Fanuc KAREL source: kd00041.KL

-- PROVISIONAL review KL for V940-1; original PC SHA256 db74242f19a3847c4d94c9fab1e78f44e8e95f5fcd8958c4a07cd94807cec2c1
-- Incomplete behavior may be omitted. Consult companion uncertainty JSON. Do not deploy.
PROGRAM KD00041
%NOLOCKGROUP
BEGIN
  -- V9_ZERO_TABLE_METADATA_HINT layout=0002_ascii; no indexed target words; source/name/runtime held
  -- UNRESOLVED_PC offsets 5-12; opcodes 9D,23
  -- UNRESOLVED_PC offsets 17-21; opcodes 7F
END KD00041
